RoboDK station: RobodkBasico-2.rdk

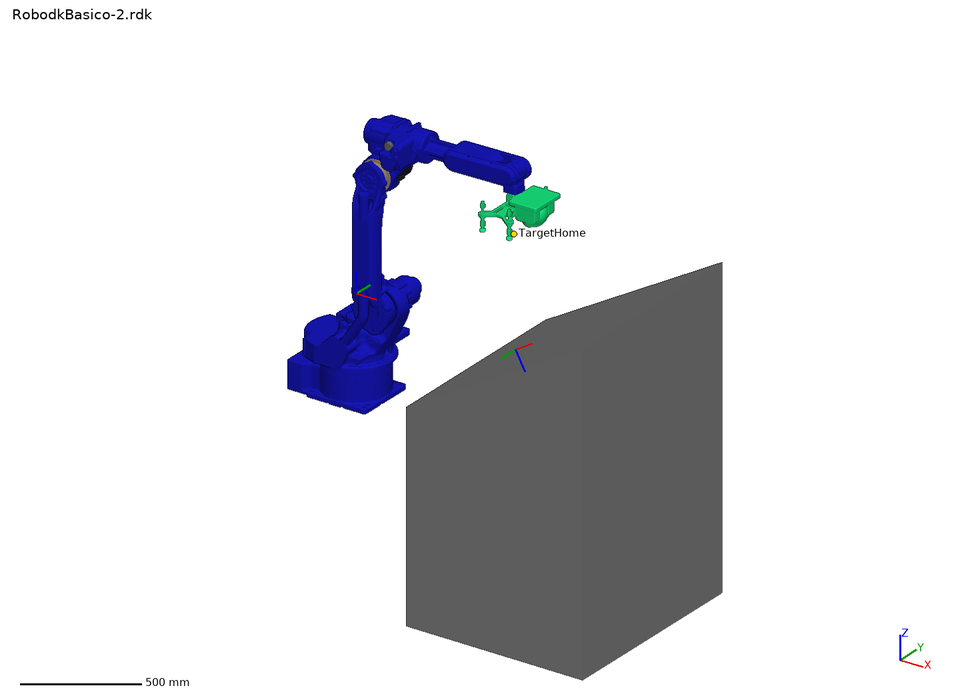
[picture v0: the station drawn from its stored meshes, robots at their saved joint values, targets as dots, program paths as lines]
Station Robodk (2) (saved by RoboDK 6.0.6). Poses are relative to the parent item; angles as X-Y-Z fixed-axis rotations.
  - frame Motoman MH6 Base at (0, 0, 450) mm
    - robot Motoman MH6: 6 axes, payload 6 kg, reach 1422 mm, repeatability 0.08 mm, weight 130 kg
        modified DH rows (alpha deg, a mm, theta deg, d mm): 0, 0, 0, 450; -90, 152, -90, 0; 0, 614, 0, 0; -90, 155, 0, 640; 90, 0, 90, 0; -90, 0, 0, 95
        base shift (0, 0, -450) mm
        joint limits [-170, -90, -175, -180, -45, -360] to [170, 155, 250, 180, 225, 360]; home [0, 0, 0, 0, 0, 0]; saved at [0, 0.258, 1.246, 0, -0.987, 0]
      - tool Ventosas, TCP at (0, 0, 190) mm, size 250 x 290 x 148 mm
    - frame Frame_from_Target1 at (823.2, -34.49, -10.13) mm, rotated rx -180 ry -30 rz 0 deg
      - target TargetHome (Cartesian target) at (225.55, -34.49, -453.06) mm, rotated rx 0 ry -30 rz 0 deg; joints [0, 0, 0, 0, 0, 0] of Motoman MH6
  - object CAJA2 at (1600, 500, 300) mm, rotated rx 180 ry 0 rz 0 deg, size 886.4 x 1000 x 1511.7 mm, geometry from CAJA2.stp
  - Python program RosPolar (listed below)
  - Python program Prog2 (listed below)

--- Python program RosPolar ---
from robodk.robolink import *    # API para comunicarte con RoboDK
from robodk.robomath import *    # Funciones matemáticas
import math

#------------------------------------------------
# 1) Conexión a RoboDK e inicialización
#------------------------------------------------
RDK = Robolink()

# Elegir un robot (si hay varios, aparece un popup)
robot = RDK.ItemUserPick("Selecciona un robot", ITEM_TYPE_ROBOT)
if not robot.Valid():
    raise Exception("No se ha seleccionado un robot válido.")



'''
# Conectar al robot físico
if not robot.Connect():
    raise Exception("No se pudo conectar al robot. Verifica que esté en modo remoto y que la configuración sea correcta.")

# Confirmar conexión
if not robot.ConnectedState():
    raise Exception("El robot no está conectado correctamente. Revisa la conexión.")

print("Robot conectado correctamente.")
'''




#------------------------------------------------
# 2) Cargar el Frame (ya existente) donde quieres dibujar
#    Ajusta el nombre si tu Frame se llama diferente
#------------------------------------------------
frame_name = "Frame_from_Target1"
frame = RDK.Item(frame_name, ITEM_TYPE_FRAME)
if not frame.Valid():
    raise Exception(f'No se encontró el Frame "{frame_name}" en la estación.')

# Asignamos este frame al robot
robot.setPoseFrame(frame)
# Usamos la herramienta activa
robot.setPoseTool(robot.PoseTool())

# Ajustes de velocidad y blending
robot.setSpeed(300)   # mm/s - Ajusta según necesites
robot.setRounding(5)  # blending (radio de curvatura)

#------------------------------------------------
# 3) Parámetros de la figura (rosa polar)
#------------------------------------------------
num_points = 720       # Cuántos puntos muestreamos (mayor = más suave)
A = 150               # Amplitud (300 mm = radio máximo)
k = 5                  # Parámetro de la rosa (pétalos). Si es impar, habrá k pétalos; si es par, 2k
z_surface = 0          # Z=0 en el plano del frame
z_safe = 50            # Altura segura para aproximarse y salir

#------------------------------------------------
# 4) Movimiento al centro en altura segura
#------------------------------------------------
# El centro de la rosa (r=0) corresponde a x=0, y=0
robot.MoveJ(transl(0, 0, z_surface - z_safe))

# Bajamos a la "superficie" (Z=0)
robot.MoveL(transl(0, 0, z_surface))

#------------------------------------------------
# 5) Dibujar la rosa polar
#    r = A * sin(k*theta)
#    x = r*cos(theta), y = r*sin(theta)
#------------------------------------------------
# Recorremos theta de 0 a 2*pi (una vuelta completa)
full_turn = 2*math.pi

for i in range(num_points+1):
    # Fracción entre 0 y 1
    t = i / num_points
    # Ángulo actual
    theta = full_turn * t

    # Calculamos r
    r = A * math.sin(k * theta)

    # Convertimos a coordenadas Cartesianas X, Y
    x = r * math.cos(theta)
    y = r * math.sin(theta)

    # Movemos linealmente (MoveL) en el plano del Frame
    robot.MoveL(transl(x, y, z_surface))

# Al terminar, subimos de nuevo para no chocar
robot.MoveL(transl(x, y, z_surface - z_safe))

print(f"¡Figura (rosa polar) completada en el frame '{frame_name}'!")

--- Python program Prog2 ---
from robodk.robolink import *
from robodk.robomath import *
import numpy as np
from matplotlib.textpath import TextPath
from matplotlib.font_manager import FontProperties

# ================= PARAMETROS =================
FRAME_NAME = "Frame_from_Target1"
Z_SURFACE = 0.0             # altura de contacto en el Frame (ajustar si el Frame esta pegado a la superficie)
Z_SAFE = 50                 # distancia positiva; al llamar se resta: Z_SURFACE - Z_SAFE
SPEED = 300                 # mm/s
ROUNDING = 0.1             # mm (menor = mas preciso, pero mas lento)

A = 150                     # tamano de la mariposa (mm)
N_SAMPLES = 50            # muestreo fino de la curva; luego RDP descarta lo redundante
TOLERANCE = 0.3             # mm de error maximo permitido al simplificar (balance puntos vs suavidad)
TEXT_W, TEXT_H = 240, 38    # caja de cada nombre (mm)
Y_NAMES = {"Felipe": -130, "Alexandra": -190}

# Orientacion de toda la composicion
MIRROR_Y = True             # corrige el efecto espejo
ROT_DEG = 90                # si sale de cabeza prueba 270; de lado prueba 0 o 180
OFFSET = np.array([300, 0])

# ================= CONEXION =================
RDK = Robolink()
robot = RDK.ItemUserPick("Selecciona un robot", ITEM_TYPE_ROBOT)
frame = RDK.Item(FRAME_NAME, ITEM_TYPE_FRAME)
home = RDK.Item("TargetHome", ITEM_TYPE_TARGET)

if not robot.Valid() or not frame.Valid() or not home.Valid():
    raise Exception(f'Falta el robot, el Frame "{FRAME_NAME}" o "TargetHome".')

'''
# Conectar al robot físico
if not robot.Connect():
    raise Exception("No se pudo conectar al robot. Verifica que esté en modo remoto y que la configuración sea correcta.")

# Confirmar conexión
state, msg = robot.ConnectedState()
if state != ROBOTCOM_READY:
    raise Exception(f"El robot no esta listo (codigo {state}): {msg}")

print("Robot conectado correctamente.")
'''

robot.setPoseFrame(frame)
robot.setPoseTool(robot.PoseTool())
robot.setSpeed(SPEED)
robot.setRounding(ROUNDING)

# ================= GEOMETRIA =================
def rdp(P, tol):
    """Ramer-Douglas-Peucker iterativo: quita puntos que desvian menos de tol mm."""
    P = np.asarray(P, dtype=float)
    keep = np.zeros(len(P), dtype=bool)
    keep[[0, -1]] = True
    stack = [(0, len(P) - 1)]
    while stack:
        i, j = stack.pop()
        if j <= i + 1:
            continue
        a, d = P[i], P[j] - P[i]
        seg = P[i + 1:j] - a
        n = np.hypot(*d)
        dist = np.hypot(*seg.T) if n == 0 else np.abs(d[0] * seg[:, 1] - d[1] * seg[:, 0]) / n
        k = np.argmax(dist)
        if dist[k] > tol:
            m = i + 1 + k
            keep[m] = True
            stack += [(i, m), (m, j)]
    return P[keep]


def transform(points):
    """Espejo en Y -> rotacion global -> traslacion."""
    a = np.radians(ROT_DEG)
    R = np.array([[np.cos(a), -np.sin(a)],
                  [np.sin(a),  np.cos(a)]])
    pts = np.asarray(points, dtype=float)
    if MIRROR_Y:
        pts = pts * [1, -1]
    return pts @ R.T + OFFSET


def butterfly():
    t = np.linspace(0, 12 * np.pi, N_SAMPLES + 1)
    r = np.exp(np.sin(t)) - 2 * np.cos(4 * t) + np.sin((2 * t - np.pi) / 24) ** 5
    r = A * r / np.max(np.abs(r))
    return rdp(np.column_stack((r * np.cos(t), r * np.sin(t))), TOLERANCE)


def text_paths(text, y_base):
    tp = TextPath((0, 0), text, size=100,
                  prop=FontProperties(family="DejaVu Sans", weight="bold"))
    polys = tp.to_polygons(closed_only=False)
    allp = np.vstack(polys)
    mn, mx = allp.min(axis=0), allp.max(axis=0)
    scale = min(TEXT_W / (mx[0] - mn[0]), TEXT_H / (mx[1] - mn[1]))
    origin = np.array([(mn[0] + mx[0]) / 2, mn[1]])   # centrado en X, base en Y
    paths = []
    for p in polys:
        p = (p - origin) * scale + [0, y_base]
        if not np.allclose(p[0], p[-1]):              # cerrar contorno
            p = np.vstack([p, p[:1]])
        paths.append(rdp(p, TOLERANCE))
    return paths


# ================= DIBUJO =================
def draw(path):
    pts = transform(path)
    x0, y0 = pts[0]
    robot.MoveJ(transl(float(x0), float(y0), Z_SURFACE - Z_SAFE))   # aproximacion
    for x, y in pts:
        robot.MoveL(transl(float(x), float(y), Z_SURFACE))          # trazo
    xf, yf = pts[-1]
    robot.MoveL(transl(float(xf), float(yf), Z_SURFACE - Z_SAFE))   # retirada


# ================= RUTINA =================
paths = [butterfly()]
for name, y in Y_NAMES.items():
    paths += text_paths(name, y)
print("Trayectorias:", len(paths), "| Puntos totales:", sum(len(p) for p in paths))

robot.MoveJ(home)          # inicio en Home
for p in paths:
    draw(p)
robot.MoveJ(home)          # final en Home
print("DIBUJO COMPLETADO")
